Fanuc KAREL source: kd00054.KL

-- PROVISIONAL review KL for V940-1; original PC SHA256 2ae57a67c7c1f6d89b14544b53996ac6c4cbf423adab7385976b28cb1768eff0
-- Incomplete behavior may be omitted. Consult companion uncertainty JSON. Do not deploy.
PROGRAM KD00054
%NOLOCKGROUP
VAR
  I : INTEGER
  J : INTEGER
  B : BOOLEAN
  R : REAL
  S : STRING[80]
BEGIN
  -- V9_ZERO_TABLE_METADATA_HINT layout=0001; no indexed target words; source/name/runtime held
  -- UNRESOLVED_PC offsets 5-28; opcodes 9D,81,18,9D,1B,9D,12,22,2E,13,04
  -- UNRESOLVED_PC offsets 33-37; opcodes 7F
END KD00054
